// TIA Portal V20 export
// export: Created 2026-10-19T18:03:06.6981204Z, ExportSetting WithDefaults, DisplayName Totally Integrated Automation Portal, DisplayVersion V20 Update 6, DisplayName TIA Portal Openness, DisplayVersion V20 Update 6, DisplayName TIA Portal Version Control Interface, DisplayVersion V20 Update 6, DisplayName SINAMICS Startdrive Advanced, DisplayVersion V20 SP1, DisplayName SINAMICS Startdrive G130, G150, S120, S150, SINAMICS MV, G220, S200, S210, DisplayVersion V20 SP1, DisplayName SINAMICS Startdrive G110M, G120, G120C, G120D, G120P, G115D, DisplayVersion V20 SP1, DisplayName STEP 7 Professional, DisplayVersion V20 Update 6, DisplayName STEP 7 Safety, DisplayVersion V20 Update 2, DisplayName WinCC Basic/Comfort/Advanced, DisplayVersion V20 Update 6, DisplayName WinCC Unified, DisplayVersion V20 Update 6
DATA_BLOCK "SB_RedAlarm"   // DB117
{ S7_Optimized_Access := 'TRUE' }
VERSION : 0.1
// stored: AutoNumber true, DBAccessibleFromOPCUA true, DBAccessibleFromWebserver true, InstanceOfName SAI_SB_RedAlert, InstanceOfType UDT, IsOnlyStoredInLoadMemory false, IsWriteProtectedInAS false
"SAI_SB_RedAlert"
   // VAR
   //    "Zero out of range" : Bool;
   //    "Symetry errors" : Bool;
   //    "LC Temperature out of normal temperature" : Bool;
   //    "Weights and measures failure" : Bool;
   //    "Foreign device detected" : Bool;
   //    "Test mode" : Bool;
   //    "LC temperature out of operatio" : Bool;
   //    "LC parameters block checksum error" : Bool;
   //    "Calibration error" : Bool;
   //    "Out of A/D range over/under" : Bool;
   //    "Checksu failure" : Bool;
   //    "Weight blocked" : Bool;
   //    "LC Missing" : Bool;
   //    "Customer-defined overload" : Bool;
   //    "Customer-defined underload" : Bool;
   // END_VAR
BEGIN
END_DATA_BLOCK
